(* IEC 61131-3 sources: plc-st-coding-agent/progress/evidence/f14_p1_20261111b/jobs/codex_deepseek-v4pro, 35 files *)

(* ---- public-easy-02.candidate_01.st ---- *)
FUNCTION_BLOCK DualWordEdgeDetector
VAR_INPUT
    value : DWORD;
END_VAR
VAR_OUTPUT
    hasChanged       : BOOL;
    hasRisingEdges   : BOOL;
    risingBits       : DWORD;
    noOfRisingBits   : USINT;
    hasFallingEdges  : BOOL;
    fallingBits      : DWORD;
    noOfFallingBits  : USINT;
END_VAR
VAR
    prevValue : DWORD;
    i : INT;
END_VAR

risingBits := value AND NOT prevValue;
fallingBits := NOT value AND prevValue;

hasRisingEdges := risingBits <> 0;
hasFallingEdges := fallingBits <> 0;
hasChanged := value <> prevValue;

noOfRisingBits := 0;
noOfFallingBits := 0;

FOR i := 0 TO 31 DO
    IF (risingBits AND SHL(DWORD#1, i)) <> 0 THEN
        noOfRisingBits := noOfRisingBits + 1;
    END_IF;

    IF (fallingBits AND SHL(DWORD#1, i)) <> 0 THEN
        noOfFallingBits := noOfFallingBits + 1;
    END_IF;
END_FOR;

prevValue := value;

(* ---- public-easy-02.candidate_02.st ---- *)
FUNCTION_BLOCK DualWordEdgeDetector
VAR_INPUT
    value : DWORD;
END_VAR
VAR_OUTPUT
    hasChanged       : BOOL;
    hasRisingEdges   : BOOL;
    risingBits       : DWORD;
    noOfRisingBits   : USINT;
    hasFallingEdges  : BOOL;
    fallingBits      : DWORD;
    noOfFallingBits  : USINT;
END_VAR
VAR
    prevValue : DWORD;
    i : INT;
END_VAR

risingBits := value AND (NOT prevValue);
fallingBits := (NOT value) AND prevValue;

hasRisingEdges := risingBits <> 0;
hasFallingEdges := fallingBits <> 0;
hasChanged := value <> prevValue;

noOfRisingBits := 0;
noOfFallingBits := 0;

FOR i := 0 TO 31 DO
    IF (risingBits AND SHL(DWORD#1, i)) <> 0 THEN
        noOfRisingBits := noOfRisingBits + 1;
    END_IF;

    IF (fallingBits AND SHL(DWORD#1, i)) <> 0 THEN
        noOfFallingBits := noOfFallingBits + 1;
    END_IF;
END_FOR;

prevValue := value;

END_FUNCTION_BLOCK

(* ---- public-easy-05.candidate_01.st ---- *)
FUNCTION_BLOCK WeldGapAlarm
VAR_INPUT
    Gap_Exceeded       : BOOL;
    Weld_E_Stop_NC     : BOOL;
    DebounceTime       : TIME;
END_VAR
VAR_OUTPUT
    Operator_Alert         : BOOL;
    Weld_Soft_Start_Active : BOOL;
END_VAR
VAR
    PowerUpTimer  : TON;
    GapTimer      : TON;
END_VAR

// 5-second power-up initialization inhibition
PowerUpTimer(IN := TRUE, PT := T#5S);
Weld_Soft_Start_Active := NOT PowerUpTimer.Q;

// Gap debounce only after initialization and while emergency stop is inactive
GapTimer(
    IN := Gap_Exceeded
          AND PowerUpTimer.Q
          AND Weld_E_Stop_NC,
    PT := DebounceTime
);

// Alarm only after full debounce, and emergency stop overrides immediately
Operator_Alert := GapTimer.Q AND Weld_E_Stop_NC;

(* ---- public-easy-05.candidate_02.st ---- *)
FUNCTION_BLOCK WeldGapAlarm
VAR_INPUT
    Gap_Exceeded       : BOOL;
    Weld_E_Stop_NC     : BOOL;
    DebounceTime       : TIME;
END_VAR
VAR_OUTPUT
    Operator_Alert         : BOOL;
    Weld_Soft_Start_Active : BOOL;
END_VAR
VAR
    PowerUpTimer  : TON;
    GapTimer      : TON;
END_VAR

PowerUpTimer(IN := TRUE, PT := T#5S);
Weld_Soft_Start_Active := NOT PowerUpTimer.Q;

GapTimer(
    IN := Gap_Exceeded
          AND PowerUpTimer.Q
          AND Weld_E_Stop_NC,
    PT := DebounceTime
);

Operator_Alert := GapTimer.Q AND Weld_E_Stop_NC;

END_FUNCTION_BLOCK

(* ---- public-easy-06.candidate_01.st ---- *)
FUNCTION_BLOCK AerationBlowerControl
VAR_INPUT
    DO_LOW : BOOL;
    AERATION_E_STOP_NC : BOOL;
END_VAR
VAR_OUTPUT
    BLOWER_RUN : BOOL;
    AERATION_BLOWER_CYCLE_COUNT : UINT;
END_VAR
VAR
    StartDelay : TON;
    BlowerRunPrev : BOOL := FALSE;
    InitDone : BOOL := FALSE;
END_VAR

IF NOT InitDone THEN
    StartDelay(IN := FALSE, PT := T#5s);
    BLOWER_RUN := FALSE;
    AERATION_BLOWER_CYCLE_COUNT := 0;
    BlowerRunPrev := FALSE;
    InitDone := TRUE;
END_IF;

StartDelay(IN := DO_LOW AND AERATION_E_STOP_NC, PT := T#5s);
BLOWER_RUN := StartDelay.Q;

IF BLOWER_RUN AND NOT BlowerRunPrev THEN
    AERATION_BLOWER_CYCLE_COUNT := AERATION_BLOWER_CYCLE_COUNT + 1;
END_IF;

BlowerRunPrev := BLOWER_RUN;
END_FUNCTION_BLOCK

(* ---- public-hard-01.candidate_01.st ---- *)
FUNCTION_BLOCK MaterialProportioningControl
VAR_INPUT
    estop            : BOOL;  (* FALSE = emergency stop active *)
    opeMode          : BOOL;  (* FALSE = manual, TRUE = automatic *)
    valveAStart      : BOOL;
    valveBStart      : BOOL;
    valveCStart      : BOOL;
    valveDStart      : BOOL;
    mixMotorStart    : BOOL;
    autoStart        : BOOL;
    processMode      : BOOL;  (* FALSE = no C, TRUE = use C until 100 cm *)
    levelSensor      : INT;   (* cm *)
    mixMotorComplete : BOOL;
END_VAR

VAR_OUTPUT
    valveARun   : BOOL;
    valveBRun   : BOOL;
    valveCRun   : BOOL;
    valveDRun   : BOOL;
    mixMotorRun : BOOL;
END_VAR

VAR
    valveAStart_RE      : BOOL;
    valveBStart_RE      : BOOL;
    valveCStart_RE      : BOOL;
    valveDStart_RE      : BOOL;
    mixMotorStart_RE    : BOOL;
    autoStart_RE        : BOOL;
    mixMotorComplete_RE : BOOL;
    modeChanged         : BOOL;

    valveAStart_prev      : BOOL;
    valveBStart_prev      : BOOL;
    valveCStart_prev      : BOOL;
    valveDStart_prev      : BOOL;
    mixMotorStart_prev    : BOOL;
    autoStart_prev        : BOOL;
    mixMotorComplete_prev : BOOL;
    opeMode_prev          : BOOL;

    manualValveA   : BOOL;
    manualValveB   : BOOL;
    manualValveC   : BOOL;
    manualValveD   : BOOL;
    manualMixMotor : BOOL;

    (* 0  = idle *)
    (* 10 = filling through valve A *)
    (* 20 = filling through valve B *)
    (* 30 = filling through valve C *)
    (* 40 = mixing *)
    (* 50 = discharging through valve D *)
    autoState : INT := 0;
END_VAR

(* Detect rising edges *)
valveAStart_RE      := valveAStart AND NOT valveAStart_prev;
valveBStart_RE      := valveBStart AND NOT valveBStart_prev;
valveCStart_RE      := valveCStart AND NOT valveCStart_prev;
valveDStart_RE      := valveDStart AND NOT valveDStart_prev;
mixMotorStart_RE    := mixMotorStart AND NOT mixMotorStart_prev;
autoStart_RE        := autoStart AND NOT autoStart_prev;
mixMotorComplete_RE := mixMotorComplete AND NOT mixMotorComplete_prev;
modeChanged         := opeMode <> opeMode_prev;

IF NOT estop THEN
    (* Emergency stop: stop everything and reset control states *)
    valveARun   := FALSE;
    valveBRun   := FALSE;
    valveCRun   := FALSE;
    valveDRun   := FALSE;
    mixMotorRun := FALSE;

    autoState      := 0;
    manualValveA   := FALSE;
    manualValveB   := FALSE;
    manualValveC   := FALSE;
    manualValveD   := FALSE;
    manualMixMotor := FALSE;

ELSIF modeChanged THEN
    (* Mode change: stop equipment and clear both control states *)
    valveARun   := FALSE;
    valveBRun   := FALSE;
    valveCRun   := FALSE;
    valveDRun   := FALSE;
    mixMotorRun := FALSE;

    autoState      := 0;
    manualValveA   := FALSE;
    manualValveB   := FALSE;
    manualValveC   := FALSE;
    manualValveD   := FALSE;
    manualMixMotor := FALSE;

ELSIF opeMode THEN
    (* Automatic mode *)

    IF autoStart_RE AND ((autoState = 0) OR (autoState = 50)) THEN
        autoState := 10;
    END_IF;

    CASE autoState OF
        10: (* Valve A is open; fill to 50 cm *)
            IF levelSensor >= 50 THEN
                autoState := 20;
            END_IF;

        20: (* Valve A closed, valve B open; fill to 80 cm *)
            IF levelSensor >= 80 THEN
                IF processMode THEN
                    autoState := 30;
                ELSE
                    autoState := 40;
                END_IF;
            END_IF;

        30: (* Valve C open; fill to 100 cm *)
            IF levelSensor >= 100 THEN
                autoState := 40;
            END_IF;

        40: (* Mixing motor running *)
            IF mixMotorComplete_RE THEN
                autoState := 50;
            END_IF;

        50: (* Valve D open; automatic process finished *)
            ;
    END_CASE;

    valveARun   := autoState = 10;
    valveBRun   := autoState = 20;
    valveCRun   := autoState = 30;
    valveDRun   := autoState = 50;
    mixMotorRun := autoState = 40;

ELSE
    (* Manual mode: each rising edge toggles the corresponding device *)
    valveARun   := manualValveA;
    valveBRun   := manualValveB;
    valveCRun   := manualValveC;
    valveDRun   := manualValveD;
    mixMotorRun := manualMixMotor;

    IF valveAStart_RE THEN
        manualValveA := NOT manualValveA;
    END_IF;

    IF valveBStart_RE THEN
        manualValveB := NOT manualValveB;
    END_IF;

    IF valveCStart_RE THEN
        manualValveC := NOT manualValveC;
    END_IF;

    IF valveDStart_RE THEN
        manualValveD := NOT manualValveD;
    END_IF;

    IF mixMotorStart_RE THEN
        manualMixMotor := NOT manualMixMotor;
    END_IF;
END_IF;

(* Store current input values for the next rising-edge detection *)
valveAStart_prev      := valveAStart;
valveBStart_prev      := valveBStart;
valveCStart_prev      := valveCStart;
valveDStart_prev      := valveDStart;
mixMotorStart_prev    := mixMotorStart;
autoStart_prev        := autoStart;
mixMotorComplete_prev := mixMotorComplete;
opeMode_prev          := opeMode;

(* ---- public-hard-01.candidate_02.st ---- *)
FUNCTION_BLOCK MaterialProportioningControl
VAR_INPUT
    estop            : BOOL;  (* FALSE: emergency stop triggered *)
    opeMode          : BOOL;  (* FALSE: manual, TRUE: automatic *)
    valveAStart      : BOOL;
    valveBStart      : BOOL;
    valveCStart      : BOOL;
    valveDStart      : BOOL;
    mixMotorStart    : BOOL;
    autoStart        : BOOL;
    processMode      : BOOL;
    levelSensor      : INT;   (* cm *)
    mixMotorComplete : BOOL;
END_VAR

VAR_OUTPUT
    valveARun   : BOOL;
    valveBRun   : BOOL;
    valveCRun   : BOOL;
    valveDRun   : BOOL;
    mixMotorRun : BOOL;
END_VAR

VAR
    valveAStart_RE      : BOOL;
    valveBStart_RE      : BOOL;
    valveCStart_RE      : BOOL;
    valveDStart_RE      : BOOL;
    mixMotorStart_RE    : BOOL;
    autoStart_RE        : BOOL;
    mixMotorComplete_RE : BOOL;
    modeChanged         : BOOL;

    valveAStart_prev      : BOOL;
    valveBStart_prev      : BOOL;
    valveCStart_prev      : BOOL;
    valveDStart_prev      : BOOL;
    mixMotorStart_prev    : BOOL;
    autoStart_prev        : BOOL;
    mixMotorComplete_prev : BOOL;
    opeMode_prev          : BOOL;

    manualValveA   : BOOL;
    manualValveB   : BOOL;
    manualValveC   : BOOL;
    manualValveD   : BOOL;
    manualMixMotor : BOOL;

    autoState : INT := 0; (* 0=idle,10=A,20=B,30=C,40=mix,50=discharge *)
END_VAR

(* Rising edge detection *)
valveAStart_RE      := valveAStart AND NOT valveAStart_prev;
valveBStart_RE      := valveBStart AND NOT valveBStart_prev;
valveCStart_RE      := valveCStart AND NOT valveCStart_prev;
valveDStart_RE      := valveDStart AND NOT valveDStart_prev;
mixMotorStart_RE    := mixMotorStart AND NOT mixMotorStart_prev;
autoStart_RE        := autoStart AND NOT autoStart_prev;
mixMotorComplete_RE := mixMotorComplete AND NOT mixMotorComplete_prev;
modeChanged         := opeMode <> opeMode_prev;

IF NOT estop THEN
    (* Emergency stop: stop all equipment and reset control states *)
    valveARun   := FALSE;
    valveBRun   := FALSE;
    valveCRun   := FALSE;
    valveDRun   := FALSE;
    mixMotorRun := FALSE;

    autoState      := 0;
    manualValveA   := FALSE;
    manualValveB   := FALSE;
    manualValveC   := FALSE;
    manualValveD   := FALSE;
    manualMixMotor := FALSE;

ELSIF modeChanged THEN
    (* Mode change: stop all equipment and clear both mode states *)
    valveARun   := FALSE;
    valveBRun   := FALSE;
    valveCRun   := FALSE;
    valveDRun   := FALSE;
    mixMotorRun := FALSE;

    autoState      := 0;
    manualValveA   := FALSE;
    manualValveB   := FALSE;
    manualValveC   := FALSE;
    manualValveD   := FALSE;
    manualMixMotor := FALSE;

ELSIF opeMode THEN
    (* Automatic mode *)
    IF autoStart_RE AND ((autoState = 0) OR (autoState = 50)) THEN
        autoState := 10;
    END_IF;

    CASE autoState OF
        10:
            IF levelSensor >= 50 THEN
                autoState := 20;
            END_IF;

        20:
            IF levelSensor >= 80 THEN
                IF processMode THEN
                    autoState := 30;
                ELSE
                    autoState := 40;
                END_IF;
            END_IF;

        30:
            IF levelSensor >= 100 THEN
                autoState := 40;
            END_IF;

        40:
            IF mixMotorComplete_RE THEN
                autoState := 50;
            END_IF;

        50:
            ; (* Valve D remains open; automatic process finished *)
    END_CASE;

    valveARun   := autoState = 10;
    valveBRun   := autoState = 20;
    valveCRun   := autoState = 30;
    valveDRun   := autoState = 50;
    mixMotorRun := autoState = 40;

ELSE
    (* Manual mode *)
    IF valveAStart_RE THEN
        manualValveA := NOT manualValveA;
    END_IF;

    IF valveBStart_RE THEN
        manualValveB := NOT manualValveB;
    END_IF;

    IF valveCStart_RE THEN
        manualValveC := NOT manualValveC;
    END_IF;

    IF valveDStart_RE THEN
        manualValveD := NOT manualValveD;
    END_IF;

    IF mixMotorStart_RE THEN
        manualMixMotor := NOT manualMixMotor;
    END_IF;

    valveARun   := manualValveA;
    valveBRun   := manualValveB;
    valveCRun   := manualValveC;
    valveDRun   := manualValveD;
    mixMotorRun := manualMixMotor;
END_IF;

(* Save current input states for next edge detection *)
valveAStart_prev      := valveAStart;
valveBStart_prev      := valveBStart;
valveCStart_prev      := valveCStart;
valveDStart_prev      := valveDStart;
mixMotorStart_prev    := mixMotorStart;
autoStart_prev        := autoStart;
mixMotorComplete_prev := mixMotorComplete;
opeMode_prev          := opeMode;

END_FUNCTION_BLOCK

(* ---- public-hard-05.candidate_01.st ---- *)
FUNCTION_BLOCK MechanicalArmControl
VAR_INPUT
    ManualMode        : BOOL;
    SingleStepMode    : BOOL;
    SingleCycleMode   : BOOL;
    ContinuousMode    : BOOL;
    EmergencyStop     : BOOL; (* FALSE: emergency stop triggered; TRUE: normal *)
    Start             : BOOL;
    DownButton        : BOOL;
    UpButton          : BOOL;
    LeftButton        : BOOL;
    RightButton       : BOOL;
    GripButton        : BOOL;
    ReleaseButton     : BOOL;
    DownLimitSwitch   : BOOL;
    UpLimitSwitch     : BOOL;
    LeftLimitSwitch   : BOOL;
    RightLimitSwitch  : BOOL;
    GripLimitSwitch   : BOOL;
    ReleaseLimitSwitch: BOOL;
END_VAR

VAR_OUTPUT
    MoveDown        : BOOL;
    MoveUp          : BOOL;
    MoveLeft        : BOOL;
    MoveRight       : BOOL;
    ActivateGrip    : BOOL;
    ActivateRelease : BOOL;
END_VAR

VAR
    StartPrev        : BOOL := FALSE;
    StartEdge        : BOOL := FALSE;
    StepActive       : BOOL := FALSE;
    StepIndex        : INT  := 0;
    SingleCycleState : INT  := 0;
    ContinuousState  : INT  := 0;
END_VAR

(* Rising edge of Start *)
StartEdge := Start AND NOT StartPrev;
StartPrev := Start;

(* Clear all commands first; emergency stop therefore disables all outputs. *)
MoveDown        := FALSE;
MoveUp          := FALSE;
MoveLeft        := FALSE;
MoveRight       := FALSE;
ActivateGrip    := FALSE;
ActivateRelease := FALSE;

IF NOT EmergencyStop THEN
    StartEdge := FALSE;

    StepActive       := FALSE;
    StepIndex        := 0;
    SingleCycleState := 0;
    ContinuousState  := 0;
ELSE
    (* ---------- Manual mode ---------- *)
    IF ManualMode THEN
        MoveDown        := DownButton    AND NOT DownLimitSwitch;
        MoveUp          := UpButton      AND NOT UpLimitSwitch;
        MoveLeft        := LeftButton    AND NOT LeftLimitSwitch;
        MoveRight       := RightButton   AND NOT RightLimitSwitch;
        ActivateGrip    := GripButton    AND NOT GripLimitSwitch;
        ActivateRelease := ReleaseButton AND NOT ReleaseLimitSwitch;
    END_IF;

    (* ---------- Single step mode ---------- *)
    IF SingleStepMode THEN
        IF StartEdge THEN
            StepIndex := StepIndex + 1;
            IF StepIndex > 8 THEN
                StepIndex := 1;
            END_IF;
            StepActive := TRUE;
        END_IF;

        IF StepActive THEN
            CASE StepIndex OF
                1: (* Down *)
                    IF DownLimitSwitch THEN
                        StepActive := FALSE;
                    ELSE
                        MoveDown := TRUE;
                    END_IF;
                2: (* Grip *)
                    IF GripLimitSwitch THEN
                        StepActive := FALSE;
                    ELSE
                        ActivateGrip := TRUE;
                    END_IF;
                3: (* Up *)
                    IF UpLimitSwitch THEN
                        StepActive := FALSE;
                    ELSE
                        MoveUp := TRUE;
                    END_IF;
                4: (* Right *)
                    IF RightLimitSwitch THEN
                        StepActive := FALSE;
                    ELSE
                        MoveRight := TRUE;
                    END_IF;
                5: (* Down *)
                    IF DownLimitSwitch THEN
                        StepActive := FALSE;
                    ELSE
                        MoveDown := TRUE;
                    END_IF;
                6: (* Release *)
                    IF ReleaseLimitSwitch THEN
                        StepActive := FALSE;
                    ELSE
                        ActivateRelease := TRUE;
                    END_IF;
                7: (* Up *)
                    IF UpLimitSwitch THEN
                        StepActive := FALSE;
                    ELSE
                        MoveUp := TRUE;
                    END_IF;
                8: (* Left *)
                    IF LeftLimitSwitch THEN
                        StepActive := FALSE;
                    ELSE
                        MoveLeft := TRUE;
                    END_IF;
            END_CASE;
        END_IF;
    ELSE
        StepActive := FALSE;
        StepIndex  := 0;
    END_IF;

    (* ---------- Single cycle mode ---------- *)
    IF SingleCycleMode THEN
        CASE SingleCycleState OF
            0: (* Idle, wait for Start *)
                IF StartEdge THEN
                    SingleCycleState := 1;
                END_IF;
            1: (* Down *)
                IF DownLimitSwitch THEN
                    SingleCycleState := 2;
                ELSE
                    MoveDown := TRUE;
                END_IF;
            2: (* Grip *)
                IF GripLimitSwitch THEN
                    SingleCycleState := 3;
                ELSE
                    ActivateGrip := TRUE;
                END_IF;
            3: (* Up *)
                IF UpLimitSwitch THEN
                    SingleCycleState := 4;
                ELSE
                    MoveUp := TRUE;
                END_IF;
            4: (* Right *)
                IF RightLimitSwitch THEN
                    SingleCycleState := 5;
                ELSE
                    MoveRight := TRUE;
                END_IF;
            5: (* Down *)
                IF DownLimitSwitch THEN
                    SingleCycleState := 6;
                ELSE
                    MoveDown := TRUE;
                END_IF;
            6: (* Release *)
                IF ReleaseLimitSwitch THEN
                    SingleCycleState := 7;
                ELSE
                    ActivateRelease := TRUE;
                END_IF;
            7: (* Up *)
                IF UpLimitSwitch THEN
                    SingleCycleState := 8;
                ELSE
                    MoveUp := TRUE;
                END_IF;
            8: (* Left *)
                IF LeftLimitSwitch THEN
                    SingleCycleState := 9;
                ELSE
                    MoveLeft := TRUE;
                END_IF;
            9: (* Completed; wait for next Start *)
                IF StartEdge THEN
                    SingleCycleState := 1;
                END_IF;
        END_CASE;
    ELSE
        SingleCycleState := 0;
    END_IF;

    (* ---------- Continuous mode ---------- *)
    IF ContinuousMode THEN
        CASE ContinuousState OF
            0: (* Idle, wait for Start *)
                IF StartEdge THEN
                    ContinuousState := 1;
                END_IF;
            1: (* Down *)
                IF DownLimitSwitch THEN
                    ContinuousState := 2;
                ELSE
                    MoveDown := TRUE;
                END_IF;
            2: (* Grip *)
                IF GripLimitSwitch THEN
                    ContinuousState := 3;
                ELSE
                    ActivateGrip := TRUE;
                END_IF;
            3: (* Up *)
                IF UpLimitSwitch THEN
                    ContinuousState := 4;
                ELSE
                    MoveUp := TRUE;
                END_IF;
            4: (* Right *)
                IF RightLimitSwitch THEN
                    ContinuousState := 5;
                ELSE
                    MoveRight := TRUE;
                END_IF;
            5: (* Down *)
                IF DownLimitSwitch THEN
                    ContinuousState := 6;
                ELSE
                    MoveDown := TRUE;
                END_IF;
            6: (* Release *)
                IF ReleaseLimitSwitch THEN
                    ContinuousState := 7;
                ELSE
                    ActivateRelease := TRUE;
                END_IF;
            7: (* Up *)
                IF UpLimitSwitch THEN
                    ContinuousState := 8;
                ELSE
                    MoveUp := TRUE;
                END_IF;
            8: (* Left, then immediately start the next cycle *)
                IF LeftLimitSwitch THEN
                    ContinuousState := 1;
                ELSE
                    MoveLeft := TRUE;
                END_IF;
        END_CASE;
    ELSE
        ContinuousState := 0;
    END_IF;
END_IF;

END_FUNCTION_BLOCK

(* ---- public-medium-01.candidate_01.st ---- *)
TYPE ST_Pump :
STRUCT
    priority  : INT;
    selection : BOOL;
    RunComd   : BOOL;
END_STRUCT
END_TYPE

FUNCTION_BLOCK FB_MultiPumpControl
VAR_INPUT
    mode  : BOOL; // FALSE: Manual, TRUE: Automatic
    start : BOOL; // Start selected pumps
    stop  : BOOL; // Stop all pumps
END_VAR
VAR_IN_OUT
    pumpGroup : ARRAY[1..5] OF ST_Pump;
END_VAR
VAR
    runActive   : BOOL := FALSE;
    selected    : ARRAY[1..5] OF BOOL;
    i           : INT;
    rank        : INT;
    bestIndex   : INT;
    bestPriority: INT;
END_VAR

IF stop THEN
    runActive := FALSE;
ELSIF start THEN
    runActive := TRUE;
END_IF;

FOR i := 1 TO 5 DO
    selected[i] := FALSE;
END_FOR;

IF runActive THEN
    IF mode THEN
        FOR rank := 1 TO 3 DO
            bestIndex := 0;
            bestPriority := 0;

            FOR i := 1 TO 5 DO
                IF NOT selected[i] THEN
                    IF (bestIndex = 0) OR (pumpGroup[i].priority > bestPriority) THEN
                        bestIndex := i;
                        bestPriority := pumpGroup[i].priority;
                    END_IF;
                END_IF;
            END_FOR;

            IF bestIndex <> 0 THEN
                selected[bestIndex] := TRUE;
            END_IF;
        END_FOR;
    ELSE
        FOR i := 1 TO 5 DO
            selected[i] := pumpGroup[i].selection;
        END_FOR;
    END_IF;
END_IF;

FOR i := 1 TO 5 DO
    pumpGroup[i].RunComd := selected[i] AND runActive;
END_FOR;

(* ---- public-medium-01.candidate_02.st ---- *)
TYPE ST_Pump :
STRUCT
    priority  : INT;
    selection : BOOL;
    RunComd   : BOOL;
END_STRUCT
END_TYPE

FUNCTION_BLOCK FB_MultiPumpControl
VAR_INPUT
    mode  : BOOL; // FALSE: Manual, TRUE: Automatic
    start : BOOL; // Start selected pumps
    stop  : BOOL; // Stop all pumps
END_VAR
VAR_IN_OUT
    pumpGroup : ARRAY[1..5] OF ST_Pump;
END_VAR
VAR
    runActive   : BOOL := FALSE;
    selected    : ARRAY[1..5] OF BOOL;
    i           : INT;
    rank        : INT;
    bestIndex   : INT;
    bestPriority: INT;
END_VAR

IF stop THEN
    runActive := FALSE;
ELSIF start THEN
    runActive := TRUE;
END_IF;

FOR i := 1 TO 5 DO
    selected[i] := FALSE;
END_FOR;

IF runActive THEN
    IF mode THEN
        FOR rank := 1 TO 3 DO
            bestIndex := 0;
            bestPriority := 0;

            FOR i := 1 TO 5 DO
                IF NOT selected[i] THEN
                    IF (bestIndex = 0) OR (pumpGroup[i].priority > bestPriority) THEN
                        bestIndex := i;
                        bestPriority := pumpGroup[i].priority;
                    END_IF;
                END_IF;
            END_FOR;

            IF bestIndex <> 0 THEN
                selected[bestIndex] := TRUE;
            END_IF;
        END_FOR;
    ELSE
        FOR i := 1 TO 5 DO
            selected[i] := pumpGroup[i].selection;
        END_FOR;
    END_IF;
END_IF;

FOR i := 1 TO 5 DO
    pumpGroup[i].RunComd := selected[i] AND runActive;
END_FOR;

END_FUNCTION_BLOCK

(* ---- public-medium-04.candidate_01.st ---- *)
FUNCTION_BLOCK FB_TemperatureControl
VAR_INPUT
    TemperatureSensorInput : REAL;
    SetTemperature : REAL;
END_VAR
VAR_OUTPUT
    CurrentTemperature : REAL;
    SetTempDisplay : REAL;
    HeaterStatus : BOOL;
    OverheatProtection : BOOL;
    HeaterOutput : BOOL;
END_VAR
VAR
    SensorFault : BOOL;
    HeaterCommand : BOOL;
    HeaterOnTimer : TON;
    CoolDownTimer : TON;
END_VAR

(* Display values *)
CurrentTemperature := TemperatureSensorInput;
SetTempDisplay := SetTemperature;

(* Sensor fault: valid measurement range is 0.0 to 100.0 *)
SensorFault := (TemperatureSensorInput < 0.0) OR (TemperatureSensorInput > 100.0);

(* Overheating protection remains active for at least 3 seconds *)
CoolDownTimer(IN := OverheatProtection, PT := T#3S);
IF CoolDownTimer.Q THEN
    OverheatProtection := FALSE;
END_IF;

(* Normal heater command *)
HeaterCommand := (NOT SensorFault)
                 AND (NOT OverheatProtection)
                 AND (TemperatureSensorInput < SetTemperature);

(* Heater running continuously for more than 5 seconds triggers protection *)
HeaterOnTimer(IN := HeaterCommand, PT := T#5S);
IF HeaterOnTimer.Q THEN
    OverheatProtection := TRUE;
END_IF;

(* Force heater off if protection is active, including the trigger moment *)
HeaterOutput := HeaterCommand AND (NOT OverheatProtection);

(* Heater status indication *)
HeaterStatus := HeaterOutput;

END_FUNCTION_BLOCK

(* ---- public-medium-06.candidate_01.st ---- *)
FUNCTION_BLOCK FB_SlabThicknessFaultMonitor
VAR_INPUT
    THICKNESS_FAULT        : BOOL;
    THICKNESS_SIGNAL_VALID : BOOL;
    CUTTING_RUN            : BOOL;
    FaultTimestamp         : DINT;
    CycleTime              : TIME; (* Must be positive *)
END_VAR
VAR_OUTPUT
    THICKNESS_ALARM        : BOOL;
    Slab_Fault_Counter     : UINT;
    Slab_Runtime_Accumulator : LTIME;
    Slab_Fault_History     : ARRAY[0..4] OF DINT; (* Read-only to callers *)
END_VAR
VAR
    Initialized    : BOOL;
    ValidFault     : BOOL;
    FaultRise      : R_TRIG;
    HoldTimer      : TON;
    HoldActive     : BOOL;
    HistoryStore   : ARRAY[0..4] OF DINT;
    i              : INT;
END_VAR

ValidFault := THICKNESS_SIGNAL_VALID AND THICKNESS_FAULT;

(* Power-up initialization *)
IF NOT Initialized THEN
    Slab_Fault_Counter := UINT#0;
    Slab_Runtime_Accumulator := LTIME#0S;

    FOR i := 0 TO 4 DO
        HistoryStore[i] := DINT#0;
    END_FOR;

    HoldActive := FALSE;
    HoldTimer(IN := FALSE, PT := T#500MS);
    Initialized := TRUE;
END_IF;

FaultRise(CLK := ValidFault);

IF NOT THICKNESS_SIGNAL_VALID THEN
    (* Signal invalid: alarm off, no holding, no fault records *)
    THICKNESS_ALARM := FALSE;
    HoldActive := FALSE;
    HoldTimer(IN := FALSE, PT := T#500MS);
ELSE
    IF FaultRise.Q THEN
        (* New valid thickness fault occurrence *)
        Slab_Fault_Counter := Slab_Fault_Counter + UINT#1;

        FOR i := 4 TO 1 BY -1 DO
            HistoryStore[i] := HistoryStore[i - 1];
        END_FOR;
        HistoryStore[0] := FaultTimestamp;

        (* Retrigger the minimum alarm hold *)
        HoldActive := FALSE;
    END_IF;

    HoldTimer(IN := HoldActive, PT := T#500MS);

    IF HoldTimer.Q THEN
        HoldActive := FALSE;
    END_IF;

    IF FaultRise.Q THEN
        HoldActive := TRUE;
    END_IF;

    THICKNESS_ALARM := THICKNESS_FAULT OR HoldActive;
END_IF;

(* Accumulate normal cutting runtime only under valid, fault-free running conditions *)
IF THICKNESS_SIGNAL_VALID
   AND CUTTING_RUN
   AND NOT THICKNESS_FAULT
   AND (CycleTime > T#0MS) THEN
    Slab_Runtime_Accumulator := Slab_Runtime_Accumulator + TIME_TO_LTIME(CycleTime);
END_IF;

(* Expose history as a copy; internal storage remains protected from direct caller changes *)
Slab_Fault_History := HistoryStore;

(* ---- public-medium-06.candidate_02.st ---- *)
FUNCTION_BLOCK FB_SlabThicknessFaultMonitor
VAR_INPUT
    THICKNESS_FAULT        : BOOL;
    THICKNESS_SIGNAL_VALID : BOOL;
    CUTTING_RUN            : BOOL;
    FaultTimestamp         : DINT;
    CycleTime              : TIME; (* Must be positive *)
END_VAR
VAR_OUTPUT
    THICKNESS_ALARM        : BOOL;
    Slab_Fault_Counter     : UINT;
    Slab_Runtime_Accumulator : LTIME;
    Slab_Fault_History     : ARRAY[0..4] OF DINT; (* Read-only to callers *)
END_VAR
VAR
    Initialized    : BOOL;
    ValidFault     : BOOL;
    FaultRise      : R_TRIG;
    HoldTimer      : TON;
    HoldActive     : BOOL;
    HistoryStore   : ARRAY[0..4] OF DINT;
    i              : INT;
END_VAR

ValidFault := THICKNESS_SIGNAL_VALID AND THICKNESS_FAULT;

(* Power-up initialization *)
IF NOT Initialized THEN
    Slab_Fault_Counter := UINT#0;
    Slab_Runtime_Accumulator := LTIME#0S;

    FOR i := 0 TO 4 DO
        HistoryStore[i] := DINT#0;
    END_FOR;

    HoldActive := FALSE;
    HoldTimer(IN := FALSE, PT := T#500MS);
    Initialized := TRUE;
END_IF;

FaultRise(CLK := ValidFault);

IF NOT THICKNESS_SIGNAL_VALID THEN
    (* Signal invalid: alarm off, no holding, no fault records *)
    THICKNESS_ALARM := FALSE;
    HoldActive := FALSE;
    HoldTimer(IN := FALSE, PT := T#500MS);
ELSE
    IF FaultRise.Q THEN
        (* New valid thickness fault occurrence *)
        Slab_Fault_Counter := Slab_Fault_Counter + UINT#1;

        FOR i := 4 TO 1 BY -1 DO
            HistoryStore[i] := HistoryStore[i - 1];
        END_FOR;
        HistoryStore[0] := FaultTimestamp;

        (* Retrigger the minimum alarm hold *)
        HoldActive := FALSE;
    END_IF;

    HoldTimer(IN := HoldActive, PT := T#500MS);

    IF HoldTimer.Q THEN
        HoldActive := FALSE;
    END_IF;

    IF FaultRise.Q THEN
        HoldActive := TRUE;
    END_IF;

    THICKNESS_ALARM := THICKNESS_FAULT OR HoldActive;
END_IF;

(* Accumulate normal cutting runtime only under valid, fault-free running conditions *)
IF THICKNESS_SIGNAL_VALID
   AND CUTTING_RUN
   AND NOT THICKNESS_FAULT
   AND (CycleTime > T#0MS) THEN
    Slab_Runtime_Accumulator := Slab_Runtime_Accumulator + TIME_TO_LTIME(CycleTime);
END_IF;

(* Expose history as a copy; internal storage remains protected from direct caller changes *)
Slab_Fault_History := HistoryStore;

END_FUNCTION_BLOCK

(* ---- public-medium-08.candidate_01.st ---- *)
FUNCTION_BLOCK IPv4Parser
VAR_INPUT
    ipText : STRING(254);
END_VAR

VAR_OUTPUT
    ipValue : UDINT;
END_VAR

VAR
    index        : DINT;
    textLen      : DINT;
    dotCount     : DINT;
    currentByte  : BYTE;
    segmentValue : UDINT;
    inSegment    : BOOL;
    segments     : ARRAY[1..4] OF UDINT;
    digitValue   : UDINT;
END_VAR

ipValue := 0;
textLen := LEN(ipText);

IF textLen = 0 THEN
    RETURN;
END_IF;

dotCount := 0;
segmentValue := 0;
inSegment := FALSE;

FOR index := 1 TO textLen DO
    currentByte := ipText[index];

    IF currentByte = 46 THEN
        IF NOT inSegment OR dotCount >= 3 THEN
            RETURN;
        END_IF;

        IF segmentValue > 255 THEN
            RETURN;
        END_IF;

        segments[dotCount + 1] := segmentValue;
        dotCount := dotCount + 1;
        segmentValue := 0;
        inSegment := FALSE;
    ELSIF currentByte >= 48 AND currentByte <= 57 THEN
        IF currentByte = 48 THEN
            digitValue := 0;
        ELSIF currentByte = 49 THEN
            digitValue := 1;
        ELSIF currentByte = 50 THEN
            digitValue := 2;
        ELSIF currentByte = 51 THEN
            digitValue := 3;
        ELSIF currentByte = 52 THEN
            digitValue := 4;
        ELSIF currentByte = 53 THEN
            digitValue := 5;
        ELSIF currentByte = 54 THEN
            digitValue := 6;
        ELSIF currentByte = 55 THEN
            digitValue := 7;
        ELSIF currentByte = 56 THEN
            digitValue := 8;
        ELSE
            digitValue := 9;
        END_IF;

        IF segmentValue > 255 THEN
            RETURN;
        END_IF;

        segmentValue := segmentValue * 10 + digitValue;

        IF segmentValue > 255 THEN
            RETURN;
        END_IF;

        inSegment := TRUE;
    ELSE
        RETURN;
    END_IF;
END_FOR;

IF NOT inSegment OR dotCount <> 3 THEN
    RETURN;
END_IF;

segments[4] := segmentValue;

ipValue := segments[1] * 16777216
         + segments[2] * 65536
         + segments[3] * 256
         + segments[4];

END_FUNCTION_BLOCK

(* ---- self-easy-01.candidate_01.st ---- *)
FUNCTION_BLOCK FB
VAR_INPUT
    enable    : BOOL;
    values    : ARRAY[1..8] OF INT;
    count     : INT;
    avgEnable : BOOL;
END_VAR
VAR_OUTPUT
    avgOut    : REAL;
END_VAR
VAR
    sumValue   : DINT;
    sampleCount: INT;
    i          : INT;
END_VAR

IF enable AND avgEnable AND (count > 0) THEN
    sampleCount := count;

    IF sampleCount > 8 THEN
        sampleCount := 8;
    END_IF;

    sumValue := 0;

    FOR i := 1 TO sampleCount BY 1 DO
        sumValue := sumValue + INT_TO_DINT(values[i]);
    END_FOR;

    avgOut := DINT_TO_REAL(sumValue) / INT_TO_REAL(sampleCount);
END_IF;

END_FUNCTION_BLOCK

(* ---- self-easy-02.candidate_01.st ---- *)
FUNCTION_BLOCK FB
VAR_INPUT
    tankLevel        : REAL;   // 储罐液位百分比 0..100
    outletFlow       : REAL;   // 出口流量 m³/h（预留观测，本题不参与逻辑）
    inletPermit      : BOOL;   // 进料许可
    resetBtn         : BOOL;   // 复位按钮，上升沿有效
END_VAR
VAR_OUTPUT
    pumpRun          : BOOL;   // 进料泵运行命令
    alarmHigh        : BOOL;   // 高液位报警，自保持
    alarmLow         : BOOL;   // 低液位报警，自保持
    outletValveOpen  : BOOL;   // 出口阀开命令
END_VAR
VAR
    prevAlarmHigh    : BOOL := FALSE;
    prevAlarmLow     : BOOL := FALSE;
    prevResetBtn     : BOOL := FALSE;
END_VAR

// 高液位报警：危险条件优先于复位沿
alarmHigh := (tankLevel >= 85.0)
             OR (prevAlarmHigh AND NOT (resetBtn AND NOT prevResetBtn));

// 低液位报警：危险条件优先于复位沿
alarmLow := (tankLevel <= 15.0)
            OR (prevAlarmLow AND NOT (resetBtn AND NOT prevResetBtn));

// 任一报警有效时禁止进料泵运行
pumpRun := inletPermit AND NOT alarmHigh AND NOT alarmLow;

// 低报警有效期间关闭出口阀，其余情况开启
outletValveOpen := NOT alarmLow;

// 保存本拍状态，供下一扫描周期使用
prevAlarmHigh := alarmHigh;
prevAlarmLow  := alarmLow;
prevResetBtn  := resetBtn;

END_FUNCTION_BLOCK

(* ---- self-hard-01.candidate_01.st ---- *)
FUNCTION_BLOCK FB
VAR_INPUT
    flowLow : BOOL;
    ackBtn : BOOL;
    sensorOK : BOOL;
END_VAR
VAR_OUTPUT
    alarmActive : BOOL;
    alarmAcked : BOOL;
    highHigh : BOOL;
END_VAR
VAR
    lastAck : BOOL;
    lastFlowLow : BOOL;
    lastAlarmActive : BOOL;
    lastAlarmAcked : BOOL;
    ackRise : BOOL;
    lastFlowAndAcked : BOOL;
    lastFlowActiveAcked : BOOL;
END_VAR

ackRise := ackBtn AND NOT lastAck;

lastFlowAndAcked := lastFlowLow AND lastAlarmAcked;
lastFlowActiveAcked := lastFlowLow AND lastAlarmActive AND lastAlarmAcked;

highHigh := NOT sensorOK;

alarmActive := flowLow OR (lastAlarmActive AND NOT ackRise AND NOT lastFlowAndAcked);
alarmAcked := alarmActive AND (NOT flowLow OR ackRise OR lastFlowActiveAcked);

lastAck := ackBtn;
lastFlowLow := flowLow;
lastAlarmActive := alarmActive;
lastAlarmAcked := alarmAcked;

END_FUNCTION_BLOCK

(* ---- self-hard-02.candidate_01.st ---- *)
FUNCTION_BLOCK FB
VAR_INPUT
    startBtn : BOOL;
    abortBtn : BOOL;
    setpoint : REAL;
    pv : REAL;
    maxDuration : INT;
END_VAR
VAR_OUTPUT
    elapsed : INT;
    phase : INT;
    timeout : BOOL;
END_VAR
VAR
    lastStartBtn : BOOL;
    startRising : BOOL;
    prevPhase : INT;
    prevElapsed : INT;
    prevTimeout : BOOL;
END_VAR

startRising := startBtn AND NOT lastStartBtn;
prevPhase := phase;
prevElapsed := elapsed;
prevTimeout := timeout;

IF abortBtn THEN
    phase := 9;
    elapsed := prevElapsed;
    timeout := prevTimeout;
ELSIF startRising THEN
    phase := 1;
    elapsed := 0;
    timeout := FALSE;
ELSIF (prevPhase = 1) OR (prevPhase = 2) THEN
    elapsed := prevElapsed + 1;

    IF maxDuration <= elapsed THEN
        timeout := TRUE;
        phase := 3;
    ELSE
        timeout := FALSE;

        IF (prevPhase = 2) OR (pv >= setpoint) THEN
            phase := 2;
        ELSE
            phase := 1;
        END_IF;
    END_IF;
ELSE
    phase := prevPhase;
    elapsed := prevElapsed;
    timeout := prevTimeout;
END_IF;

lastStartBtn := startBtn;
END_FUNCTION_BLOCK

(* ---- self-hard-03.candidate_01.st ---- *)
FUNCTION_BLOCK FB
VAR_INPUT
    pushEn : BOOL;
    pushItem : INT;
    popEn : BOOL;
END_VAR
VAR_IN_OUT
    fifo : ARRAY[1..8] OF INT;
END_VAR
VAR_OUTPUT
    count : INT := 0;
    full : BOOL := FALSE;
    empty : BOOL := TRUE;
    head : INT := 0;
END_VAR
VAR
    pushRise : BOOL;
    popRise : BOOL;
    pushPrev : BOOL := FALSE;
    popPrev : BOOL := FALSE;
    workingCount : INT;
    idx : INT;
END_VAR

pushRise := pushEn AND NOT pushPrev;
popRise := popEn AND NOT popPrev;

workingCount := count;

IF popRise AND (workingCount > 0) THEN
    IF workingCount > 1 THEN
        FOR idx := 1 TO workingCount - 1 DO
            fifo[idx] := fifo[idx + 1];
        END_FOR;
    END_IF;
    fifo[workingCount] := 0;
    workingCount := workingCount - 1;
END_IF;

IF pushRise AND (workingCount < 8) THEN
    fifo[workingCount + 1] := pushItem;
    workingCount := workingCount + 1;
END_IF;

count := workingCount;
full := (workingCount = 8);
empty := (workingCount = 0);

IF workingCount > 0 THEN
    head := fifo[1];
ELSE
    head := 0;
END_IF;

pushPrev := pushEn;
popPrev := popEn;
END_FUNCTION_BLOCK

(* ---- self-hard-04.candidate_01.st ---- *)
FUNCTION_BLOCK FB
VAR_INPUT
    demand : INT;
    runHours : ARRAY[1..5] OF LINT;
    rotated : BOOL;
END_VAR
VAR_OUTPUT
    leadPump : INT;
    lagPump : INT;
    runningCount : INT;
END_VAR
VAR
    previousLeadPump : INT := 0;
    previousLagPump : INT := 0;
    previousRunningCount : INT := 0;
    clippedDemand : INT;
    minimumPump : INT;
    minimumHours : LINT;
    lagCandidate : INT;
    pumpIndex : INT;
END_VAR

clippedDemand := demand;
IF clippedDemand < 0 THEN
    clippedDemand := 0;
ELSIF clippedDemand > 5 THEN
    clippedDemand := 5;
END_IF;

runningCount := clippedDemand;

IF clippedDemand <= 0 THEN
    leadPump := 0;
    lagPump := 0;
ELSE
    minimumHours := runHours[1];
    minimumPump := 1;
    FOR pumpIndex := 2 TO 5 DO
        IF (runHours[pumpIndex] < minimumHours) OR
           ((runHours[pumpIndex] = minimumHours) AND (pumpIndex < minimumPump)) THEN
            minimumHours := runHours[pumpIndex];
            minimumPump := pumpIndex;
        END_IF;
    END_FOR;

    IF (previousLeadPump < 1) OR (previousLeadPump > 5) THEN
        leadPump := minimumPump;
    ELSIF rotated AND
          (previousLeadPump >= 1) AND
          (previousLeadPump <= 5) AND
          (runHours[previousLeadPump] - minimumHours > 50) THEN
        leadPump := minimumPump;
    ELSE
        leadPump := previousLeadPump;
    END_IF;

    IF clippedDemand >= 2 THEN
        IF (leadPump <> previousLeadPump) OR (runningCount > previousRunningCount) THEN
            lagCandidate := 0;
            FOR pumpIndex := 1 TO 5 DO
                IF pumpIndex <> leadPump THEN
                    IF lagCandidate = 0 THEN
                        lagCandidate := pumpIndex;
                    ELSIF (runHours[pumpIndex] < runHours[lagCandidate]) OR
                          ((runHours[pumpIndex] = runHours[lagCandidate]) AND
                           (pumpIndex < lagCandidate)) THEN
                        lagCandidate := pumpIndex;
                    END_IF;
                END_IF;
            END_FOR;
            lagPump := lagCandidate;
        ELSE
            lagPump := previousLagPump;
        END_IF;
    ELSE
        lagPump := 0;
    END_IF;
END_IF;

previousLeadPump := leadPump;
previousLagPump := lagPump;
previousRunningCount := runningCount;
END_FUNCTION_BLOCK

(* ---- self-hard-05.candidate_01.st ---- *)
FUNCTION_BLOCK FB
VAR_INPUT
    runRequest : BOOL;
    flameOK : BOOL;
    o2Valid : BOOL;
    o2PV : REAL;
    baseAir : REAL;
    resetBtn : BOOL;
END_VAR
VAR_OUTPUT
    fuelPermit : BOOL;
    trimEnable : BOOL;
    airTrim : REAL;
    airCommand : REAL;
    tripLatched : BOOL;
    o2Fault : BOOL;
END_VAR
VAR
    tripMemory : BOOL;
    resetPrev : BOOL;
    resetRising : BOOL;
END_VAR

resetRising := resetBtn AND NOT resetPrev;

tripMemory := (runRequest AND NOT flameOK)
              OR (tripMemory AND NOT (resetRising AND NOT runRequest AND NOT flameOK));
tripLatched := tripMemory;

fuelPermit := runRequest AND flameOK AND NOT tripLatched;

o2Fault := NOT o2Valid OR o2PV < 0.0 OR o2PV > 21.0;

trimEnable := fuelPermit AND NOT o2Fault;

IF trimEnable THEN
    airTrim := 2.0 * (2.0 - o2PV);
    IF airTrim > 10.0 THEN
        airTrim := 10.0;
    END_IF;
    IF airTrim < -10.0 THEN
        airTrim := -10.0;
    END_IF;
ELSE
    airTrim := 0.0;
END_IF;

IF fuelPermit THEN
    airCommand := baseAir + airTrim;
    IF airCommand > 100.0 THEN
        airCommand := 100.0;
    END_IF;
    IF airCommand < 0.0 THEN
        airCommand := 0.0;
    END_IF;
ELSE
    airCommand := 0.0;
END_IF;

resetPrev := resetBtn;

(* ---- self-hard-05.candidate_02.st ---- *)
FUNCTION_BLOCK FB
VAR_INPUT
    runRequest : BOOL;
    flameOK : BOOL;
    o2Valid : BOOL;
    o2PV : REAL;
    baseAir : REAL;
    resetBtn : BOOL;
END_VAR
VAR_OUTPUT
    fuelPermit : BOOL;
    trimEnable : BOOL;
    airTrim : REAL;
    airCommand : REAL;
    tripLatched : BOOL;
    o2Fault : BOOL;
END_VAR
VAR
    tripMemory : BOOL;
    resetPrev : BOOL;
    resetRising : BOOL;
END_VAR

resetRising := resetBtn AND NOT resetPrev;

tripMemory := (runRequest AND NOT flameOK)
              OR (tripMemory AND NOT (resetRising AND NOT runRequest AND NOT flameOK));
tripLatched := tripMemory;

fuelPermit := runRequest AND flameOK AND NOT tripLatched;

o2Fault := NOT o2Valid OR o2PV < 0.0 OR o2PV > 21.0;

trimEnable := fuelPermit AND NOT o2Fault;

IF trimEnable THEN
    airTrim := 2.0 * (2.0 - o2PV);

    IF airTrim > 10.0 THEN
        airTrim := 10.0;
    END_IF;

    IF airTrim < -10.0 THEN
        airTrim := -10.0;
    END_IF;
ELSE
    airTrim := 0.0;
END_IF;

IF fuelPermit THEN
    airCommand := baseAir + airTrim;

    IF airCommand > 100.0 THEN
        airCommand := 100.0;
    END_IF;

    IF airCommand < 0.0 THEN
        airCommand := 0.0;
    END_IF;
ELSE
    airCommand := 0.0;
END_IF;

resetPrev := resetBtn;

END_FUNCTION_BLOCK

(* ---- self-hard-06.candidate_01.st ---- *)
FUNCTION_BLOCK FB
VAR_INPUT
    runRequest : BOOL;
    pressure : REAL;
    pressureValid : BOOL;
    fuelFlow : REAL;
    steamFlow : REAL;
    outletCmd : INT;
    outletFeedback : INT;
    resetBtn : BOOL;
END_VAR
VAR_OUTPUT
    tripLatched : BOOL;
    fuelPermit : BOOL;
    currentCauseMask : WORD;
    latchedCauseMask : WORD;
    diagnosticActive : BOOL;
END_VAR
VAR
    resetPrev : BOOL := FALSE;
    resetRising : BOOL;
    resetAllowed : BOOL;
    tripPending : BOOL;
    overpressureActive : BOOL;
    valveStuckActive : BOOL;
    stuckCounter : INT := 0;
END_VAR

resetRising := resetBtn AND NOT resetPrev;

overpressureActive := runRequest AND pressureValid AND (pressure >= 4500.0);

IF overpressureActive AND (outletCmd >= 50) AND (outletFeedback <= 10) THEN
    IF stuckCounter < 3 THEN
        stuckCounter := stuckCounter + 1;
    END_IF;
ELSE
    stuckCounter := 0;
END_IF;

valveStuckActive := stuckCounter >= 3;

currentCauseMask := WORD#0;

IF runRequest AND NOT pressureValid THEN
    currentCauseMask := WORD#1;
ELSIF overpressureActive THEN
    IF valveStuckActive THEN
        currentCauseMask := currentCauseMask OR WORD#2;
    END_IF;

    IF (fuelFlow >= 4.0) AND (steamFlow <= 10.0) THEN
        currentCauseMask := currentCauseMask OR WORD#4;
    END_IF;

    IF currentCauseMask = WORD#0 THEN
        currentCauseMask := WORD#8;
    END_IF;
END_IF;

resetAllowed := resetRising AND NOT runRequest AND pressureValid AND (pressure <= 4200.0);
tripPending := runRequest AND ((NOT pressureValid) OR (pressure >= 4500.0));

IF resetAllowed THEN
    tripLatched := FALSE;
ELSE
    tripLatched := tripLatched OR tripPending;
END_IF;

fuelPermit := runRequest AND NOT tripLatched;
diagnosticActive := currentCauseMask <> WORD#0;

IF tripLatched THEN
    latchedCauseMask := latchedCauseMask OR currentCauseMask;
ELSE
    latchedCauseMask := WORD#0;
END_IF;

resetPrev := resetBtn;
END_FUNCTION_BLOCK

(* ---- self-hard-07.candidate_01.st ---- *)
FUNCTION_BLOCK FB
VAR_INPUT
    mode : INT;
    resetBtn : BOOL;
    scanSeconds : REAL;
    tempSP : REAL;
    tempPV : REAL;
    flowPV : REAL;
    manualFlowSP : REAL;
    manualValve : REAL;
END_VAR

VAR_OUTPUT
    flowSP : REAL;
    valveCommand : REAL;
    fault : BOOL;
    normalMode : BOOL;
END_VAR

VAR
    firstScan : BOOL := TRUE;
    prevMode : INT := 0;
    prevResetBtn : BOOL := FALSE;
    prevFlowSP : REAL := 0.0;
    prevValveCommand : REAL := 0.0;
    prevET : REAL := 0.0;
    prevEF : REAL := 0.0;
    resetRising : BOOL;
    modeChanged : BOOL;
    eT : REAL;
    eF : REAL;
END_VAR

    fault := (mode < 0) OR (mode > 2) OR (scanSeconds <= 0.0) OR (scanSeconds > 10.0);
    resetRising := resetBtn AND NOT prevResetBtn;
    modeChanged := (NOT firstScan) AND (mode <> prevMode);
    normalMode := (NOT firstScan) AND (mode = prevMode) AND (NOT fault) AND (NOT resetRising);

    eT := tempSP - tempPV;

    IF fault THEN
        flowSP := manualFlowSP;
        valveCommand := manualValve;
    ELSIF firstScan THEN
        flowSP := manualFlowSP;
        valveCommand := manualValve;
    ELSIF resetRising THEN
        flowSP := manualFlowSP;
        valveCommand := manualValve;
    ELSIF modeChanged THEN
        IF mode = 2 THEN
            flowSP := prevFlowSP;
            valveCommand := prevValveCommand;
        ELSE
            flowSP := manualFlowSP;
            valveCommand := prevValveCommand;
        END_IF;
    ELSE
        CASE mode OF
            0:
                flowSP := manualFlowSP;
                valveCommand := manualValve;

            1:
                flowSP := manualFlowSP;
                eF := flowSP - flowPV;
                valveCommand := LIMIT(0.0,
                    2.0 * eF + ((prevValveCommand - 2.0 * prevEF) + 0.5 * eF * scanSeconds),
                    100.0);

            2:
                flowSP := LIMIT(0.0,
                    1.0 * eT + ((prevFlowSP - 1.0 * prevET) + 0.2 * eT * scanSeconds),
                    50.0);
                eF := flowSP - flowPV;
                valveCommand := LIMIT(0.0,
                    2.0 * eF + ((prevValveCommand - 2.0 * prevEF) + 0.5 * eF * scanSeconds),
                    100.0);

            ELSE
                flowSP := manualFlowSP;
                valveCommand := manualValve;
        END_CASE;
    END_IF;

    prevResetBtn := resetBtn;
    prevMode := mode;
    prevFlowSP := flowSP;
    prevValveCommand := valveCommand;
    prevET := eT;
    prevEF := flowSP - flowPV;
    firstScan := FALSE;
END_FUNCTION_BLOCK

(* ---- self-medium-01.candidate_01.st ---- *)
FUNCTION_BLOCK FB
VAR_INPUT
    recipe : ARRAY[1..8] OF ST_Recipe;
    selSlot : INT;
    loadCmd : BOOL;
    running : BOOL;
END_VAR
VAR_OUTPUT
    valid : BOOL;
    loadedID : INT;
END_VAR
VAR
    previousLoadCmd : BOOL := FALSE;
    previousValid : BOOL := FALSE;
    previousLoadedID : INT := 0;
    loadEdge : BOOL;
    slotInRange : BOOL;
    slotNonEmpty : BOOL;
    ratioInRange : BOOL;
    temperatureInRange : BOOL;
END_VAR

loadEdge := loadCmd AND NOT previousLoadCmd;

loadedID := previousLoadedID;
valid := previousValid;

IF loadEdge AND NOT running THEN
    slotInRange := (selSlot >= 1) AND (selSlot <= 8);

    IF slotInRange THEN
        slotNonEmpty := recipe[selSlot].recipeID <> 0;
        ratioInRange := (recipe[selSlot].totalRatio >= 99.0)
                        AND (recipe[selSlot].totalRatio <= 101.0);
        temperatureInRange := (recipe[selSlot].temperature >= 30.0)
                              AND (recipe[selSlot].temperature <= 180.0);

        IF slotNonEmpty AND ratioInRange AND temperatureInRange THEN
            valid := TRUE;
            loadedID := recipe[selSlot].recipeID;
        ELSE
            valid := FALSE;
            loadedID := 0;
        END_IF;
    ELSE
        valid := FALSE;
        loadedID := 0;
    END_IF;
END_IF;

previousLoadCmd := loadCmd;
previousValid := valid;
previousLoadedID := loadedID;

(* ---- self-medium-01.candidate_02.st ---- *)
TYPE ST_Recipe :
STRUCT
    recipeID : INT;
    totalRatio : REAL;
    temperature : REAL;
END_STRUCT
END_TYPE

FUNCTION_BLOCK FB
VAR_INPUT
    recipe : ARRAY[1..8] OF ST_Recipe;
    selSlot : INT;
    loadCmd : BOOL;
    running : BOOL;
END_VAR
VAR_OUTPUT
    valid : BOOL;
    loadedID : INT;
END_VAR
VAR
    previousLoadCmd : BOOL := FALSE;
    previousValid : BOOL := FALSE;
    previousLoadedID : INT := 0;
    loadEdge : BOOL;
    slotInRange : BOOL;
    slotNonEmpty : BOOL;
    ratioInRange : BOOL;
    temperatureInRange : BOOL;
END_VAR

loadEdge := loadCmd AND NOT previousLoadCmd;

loadedID := previousLoadedID;
valid := previousValid;

IF loadEdge AND NOT running THEN
    slotInRange := (selSlot >= 1) AND (selSlot <= 8);

    IF slotInRange THEN
        slotNonEmpty := recipe[selSlot].recipeID <> 0;
        ratioInRange := (recipe[selSlot].totalRatio >= 99.0)
                        AND (recipe[selSlot].totalRatio <= 101.0);
        temperatureInRange := (recipe[selSlot].temperature >= 30.0)
                              AND (recipe[selSlot].temperature <= 180.0);

        IF slotNonEmpty AND ratioInRange AND temperatureInRange THEN
            valid := TRUE;
            loadedID := recipe[selSlot].recipeID;
        ELSE
            valid := FALSE;
            loadedID := 0;
        END_IF;
    ELSE
        valid := FALSE;
        loadedID := 0;
    END_IF;
END_IF;

previousLoadCmd := loadCmd;
previousValid := valid;
previousLoadedID := loadedID;

END_FUNCTION_BLOCK

(* ---- self-medium-02.candidate_01.st ---- *)
FUNCTION_BLOCK FB
VAR_INPUT
    enable : BOOL;
    rawValue : REAL;
END_VAR
VAR_OUTPUT
    filteredValue : REAL;
    windowFull : BOOL;
    sampleCount : INT;
END_VAR
VAR
    buffer : ARRAY[0..7] OF REAL;
    writeIndex : INT := 0;
    validCount : INT := 0;
    sum : REAL;
    loopIndex : INT;
END_VAR

IF enable THEN
    buffer[writeIndex] := rawValue;
    writeIndex := (writeIndex + 1) MOD 8;

    IF validCount < 8 THEN
        validCount := validCount + 1;
    END_IF;

    IF validCount = 1 THEN
        filteredValue := rawValue;
    ELSIF validCount = 2 THEN
        filteredValue := (buffer[0] + buffer[1]) / 2.0;
    ELSE
        sum := 0.0;
        FOR loopIndex := 0 TO validCount - 1 DO
            sum := sum + buffer[loopIndex];
        END_FOR;
        filteredValue := sum / INT_TO_REAL(validCount);
    END_IF;

    sampleCount := validCount;
    windowFull := validCount >= 8;
ELSE
    FOR loopIndex := 0 TO 7 DO
        buffer[loopIndex] := 0.0;
    END_FOR;

    writeIndex := 0;
    validCount := 0;
    sampleCount := 0;
    windowFull := FALSE;
END_IF

(* ---- self-medium-02.candidate_02.st ---- *)
FUNCTION_BLOCK FB
VAR_INPUT
    enable : BOOL;
    rawValue : REAL;
END_VAR
VAR_OUTPUT
    filteredValue : REAL;
    windowFull : BOOL;
    sampleCount : INT;
END_VAR
VAR
    buffer : ARRAY[0..7] OF REAL;
    writeIndex : INT := 0;
    validCount : INT := 0;
    sum : REAL;
    loopIndex : INT;
END_VAR

IF enable THEN
    buffer[writeIndex] := rawValue;
    writeIndex := (writeIndex + 1) MOD 8;

    IF validCount < 8 THEN
        validCount := validCount + 1;
    END_IF;

    IF validCount = 1 THEN
        filteredValue := rawValue;
    ELSIF validCount = 2 THEN
        filteredValue := (buffer[0] + buffer[1]) / 2.0;
    ELSE
        sum := 0.0;
        FOR loopIndex := 0 TO validCount - 1 DO
            sum := sum + buffer[loopIndex];
        END_FOR;
        filteredValue := sum / INT_TO_REAL(validCount);
    END_IF;

    sampleCount := validCount;
    windowFull := validCount >= 8;
ELSE
    FOR loopIndex := 0 TO 7 DO
        buffer[loopIndex] := 0.0;
    END_FOR;

    writeIndex := 0;
    validCount := 0;
    sampleCount := 0;
    windowFull := FALSE;
END_IF
END_FUNCTION_BLOCK

(* ---- self-medium-03.candidate_01.st ---- *)
FUNCTION_BLOCK FB
VAR_INPUT
    openBtn    : BOOL;
    closeBtn   : BOOL;
    openLimit  : BOOL;
    closeLimit : BOOL;
    obstacle   : BOOL;
END_VAR
VAR_OUTPUT
    motorUp    : BOOL;
    motorDown  : BOOL;
    errorFlag  : BOOL;
END_VAR
VAR
    state         : INT := 0; (* 0=IDLE, 1=OPENING, 2=CLOSING, 3=FAULT *)
    prevOpenBtn   : BOOL := FALSE;
    prevCloseBtn  : BOOL := FALSE;
    prevObstacle  : BOOL := FALSE;
    prevMotorUp   : BOOL := FALSE;
    prevMotorDown : BOOL := FALSE;
    prevErrorFlag : BOOL := FALSE;
END_VAR

VAR
    openRising  : BOOL;
    closeRising : BOOL;
    comboRising : BOOL;
END_VAR

openRising  := openBtn AND NOT prevOpenBtn;
closeRising := closeBtn AND NOT prevCloseBtn;
comboRising := (openBtn AND closeBtn) AND NOT (prevOpenBtn AND prevCloseBtn);

IF obstacle THEN
    state := 3;
    motorUp := FALSE;
    motorDown := FALSE;
    errorFlag := TRUE;
ELSIF state = 3 THEN
    motorUp := FALSE;
    motorDown := FALSE;
    IF comboRising THEN
        state := 0;
        errorFlag := FALSE;
    ELSE
        errorFlag := TRUE;
    END_IF;
ELSIF state = 1 THEN
    errorFlag := FALSE;
    motorDown := FALSE;
    IF openLimit THEN
        motorUp := FALSE;
        state := 0;
    ELSE
        motorUp := TRUE;
    END_IF;
ELSIF state = 2 THEN
    errorFlag := FALSE;
    motorUp := FALSE;
    IF closeLimit THEN
        motorDown := FALSE;
        state := 0;
    ELSE
        motorDown := TRUE;
    END_IF;
ELSE (* state = 0: IDLE *)
    motorUp := FALSE;
    motorDown := FALSE;
    errorFlag := FALSE;

    IF openRising AND NOT closeBtn AND NOT openLimit THEN
        motorUp := TRUE;
        state := 1;
    ELSIF closeRising AND NOT openBtn AND NOT closeLimit THEN
        motorDown := TRUE;
        state := 2;
    END_IF;
END_IF;

prevOpenBtn   := openBtn;
prevCloseBtn  := closeBtn;
prevObstacle  := obstacle;
prevMotorUp   := motorUp;
prevMotorDown := motorDown;
prevErrorFlag := errorFlag;
END_FUNCTION_BLOCK

(* ---- self-medium-04.candidate_01.st ---- *)
FUNCTION_BLOCK FB
VAR_INPUT
    startBtn : BOOL;
    resetBtn : BOOL;
    doneSensor : BOOL;
    targetVol : REAL;
    flowVol : REAL;
END_VAR
VAR_OUTPUT
    valveOpen : BOOL;
    fillsToday : INT;
END_VAR
VAR
    prevStartBtn : BOOL;
    prevResetBtn : BOOL;
    prevValveOpen : BOOL;
    bottleVol : REAL;
    pendingConfirm : BOOL;
    valveState : BOOL;
    fillCount : INT;
END_VAR

IF resetBtn AND NOT prevResetBtn THEN
    fillCount := 0;
    bottleVol := 0.0;
    valveState := FALSE;
    pendingConfirm := FALSE;
ELSE
    IF startBtn AND NOT prevStartBtn THEN
        IF NOT prevValveOpen THEN
            pendingConfirm := FALSE;
            bottleVol := 0.0;
            valveState := TRUE;
        END_IF;
    END_IF;

    IF valveState THEN
        bottleVol := bottleVol + flowVol;
        IF bottleVol >= targetVol THEN
            valveState := FALSE;
            pendingConfirm := TRUE;
        END_IF;
    END_IF;

    IF doneSensor AND pendingConfirm AND NOT valveState THEN
        IF fillCount < 32767 THEN
            fillCount := fillCount + 1;
        END_IF;
        pendingConfirm := FALSE;
    END_IF;
END_IF;

valveOpen := valveState;
fillsToday := fillCount;

prevStartBtn := startBtn;
prevResetBtn := resetBtn;
prevValveOpen := valveState;

(* ---- self-medium-04.candidate_02.st ---- *)
FUNCTION_BLOCK FB
VAR_INPUT
    startBtn : BOOL;
    resetBtn : BOOL;
    doneSensor : BOOL;
    targetVol : REAL;
    flowVol : REAL;
END_VAR
VAR_OUTPUT
    valveOpen : BOOL;
    fillsToday : INT;
END_VAR
VAR
    prevStartBtn : BOOL;
    prevResetBtn : BOOL;
    prevValveOpen : BOOL;
    bottleVol : REAL;
    pendingConfirm : BOOL;
    valveState : BOOL;
    fillCount : INT;
END_VAR

IF resetBtn AND NOT prevResetBtn THEN
    fillCount := 0;
    bottleVol := 0.0;
    valveState := FALSE;
    pendingConfirm := FALSE;
ELSE
    IF startBtn AND NOT prevStartBtn THEN
        IF NOT prevValveOpen THEN
            pendingConfirm := FALSE;
            bottleVol := 0.0;
            valveState := TRUE;
        END_IF;
    END_IF;

    IF valveState THEN
        bottleVol := bottleVol + flowVol;
        IF bottleVol >= targetVol THEN
            valveState := FALSE;
            pendingConfirm := TRUE;
        END_IF;
    END_IF;

    IF doneSensor AND pendingConfirm AND NOT valveState THEN
        IF fillCount < 32767 THEN
            fillCount := fillCount + 1;
        END_IF;
        pendingConfirm := FALSE;
    END_IF;
END_IF;

valveOpen := valveState;
fillsToday := fillCount;

prevStartBtn := startBtn;
prevResetBtn := resetBtn;
prevValveOpen := valveState;

END_FUNCTION_BLOCK

(* ---- self-medium-05.candidate_01.st ---- *)
FUNCTION_BLOCK FB
VAR_INPUT
    enable : BOOL;
    resetBtn : BOOL;
    scanSeconds : LREAL;
    steamFlow : LREAL;
    fuelFlow : LREAL;
    steamTemp : LREAL;
    steamPressure : LREAL;
END_VAR
VAR_OUTPUT
    qualified : BOOL;
    dataFault : BOOL;
    qualifiedTon : LREAL;
    fuelTon : LREAL;
    revenue : LREAL;
    cost : LREAL;
    netProfit : LREAL;
END_VAR
VAR
    resetBtnPrev : BOOL;
END_VAR

qualified := (steamTemp >= 447.0)
             AND (steamTemp <= 453.0)
             AND (steamPressure >= 3750.0)
             AND (steamPressure <= 3850.0);

dataFault := (scanSeconds <= 0.0)
             OR (scanSeconds > 10.0)
             OR (steamFlow < 0.0)
             OR (steamFlow > 90.0)
             OR (fuelFlow < 0.0)
             OR (fuelFlow > 6.0);

IF resetBtn AND NOT resetBtnPrev THEN
    qualifiedTon := 0.0;
    fuelTon := 0.0;
ELSIF dataFault THEN
    qualifiedTon := qualifiedTon;
    fuelTon := fuelTon;
ELSIF enable THEN
    fuelTon := fuelTon + fuelFlow * scanSeconds / 1000.0;

    IF qualified THEN
        qualifiedTon := qualifiedTon + steamFlow * scanSeconds / 1000.0;
    END_IF;
ELSIF NOT enable THEN
    qualifiedTon := qualifiedTon;
    fuelTon := fuelTon;
END_IF;

revenue := qualifiedTon * 280.0;
cost := fuelTon * 1500.0;
netProfit := revenue - cost;

resetBtnPrev := resetBtn;

(* ---- self-medium-05.candidate_02.st ---- *)
FUNCTION_BLOCK FB
VAR_INPUT
    enable : BOOL;
    resetBtn : BOOL;
    scanSeconds : LREAL;
    steamFlow : LREAL;
    fuelFlow : LREAL;
    steamTemp : LREAL;
    steamPressure : LREAL;
END_VAR
VAR_OUTPUT
    qualified : BOOL;
    dataFault : BOOL;
    qualifiedTon : LREAL;
    fuelTon : LREAL;
    revenue : LREAL;
    cost : LREAL;
    netProfit : LREAL;
END_VAR
VAR
    resetBtnPrev : BOOL := FALSE;
    qualifiedAcc : LREAL := 0.0;
    fuelAcc : LREAL := 0.0;
END_VAR

qualified := (steamTemp >= 447.0)
             AND (steamTemp <= 453.0)
             AND (steamPressure >= 3750.0)
             AND (steamPressure <= 3850.0);

dataFault := (scanSeconds <= 0.0)
             OR (scanSeconds > 10.0)
             OR (steamFlow < 0.0)
             OR (steamFlow > 90.0)
             OR (fuelFlow < 0.0)
             OR (fuelFlow > 6.0);

IF resetBtn AND NOT resetBtnPrev THEN
    qualifiedAcc := 0.0;
    fuelAcc := 0.0;
ELSE
    IF enable AND NOT dataFault THEN
        fuelAcc := fuelAcc + fuelFlow * scanSeconds / 1000.0;

        IF qualified THEN
            qualifiedAcc := qualifiedAcc + steamFlow * scanSeconds / 1000.0;
        END_IF;
    END_IF;
END_IF;

qualifiedTon := qualifiedAcc;
fuelTon := fuelAcc;

revenue := qualifiedTon * 280.0;
cost := fuelTon * 1500.0;
netProfit := revenue - cost;

resetBtnPrev := resetBtn;

END_FUNCTION_BLOCK

(* ---- public-easy-01.candidate_01.st ---- *)
PROGRAM FillingLineControl
VAR_INPUT
    bottleSensor : BOOL;
    cleaningConfirmButton : BOOL;
    fillingConfirmButton : BOOL;
    cappingConfirmButton : BOOL;
    packingConfirmButton : BOOL;
    finishedButton : BOOL;
END_VAR
VAR_OUTPUT
    Pump_Motor : BOOL;
    Filling_Valve : BOOL;
    Capping_Machine : BOOL;
    Packing_Machine : BOOL;
    Completion_Light : BOOL;
END_VAR
VAR
    State : INT := 0;
    bottleSensorR : R_TRIG;
    cleaningConfirmR : R_TRIG;
    fillingConfirmR : R_TRIG;
    cappingConfirmR : R_TRIG;
    packingConfirmR : R_TRIG;
    finishedR : R_TRIG;
END_VAR

bottleSensorR(CLK := bottleSensor);
cleaningConfirmR(CLK := cleaningConfirmButton);
fillingConfirmR(CLK := fillingConfirmButton);
cappingConfirmR(CLK := cappingConfirmButton);
packingConfirmR(CLK := packingConfirmButton);
finishedR(CLK := finishedButton);

Pump_Motor := FALSE;
Filling_Valve := FALSE;
Capping_Machine := FALSE;
Packing_Machine := FALSE;
Completion_Light := FALSE;

CASE State OF
    1:
        Pump_Motor := TRUE;
    2:
        Filling_Valve := TRUE;
    3:
        Capping_Machine := TRUE;
    4:
        Packing_Machine := TRUE;
    5:
        Completion_Light := TRUE;
END_CASE

IF State = 0 AND bottleSensorR.Q THEN
    State := 1;
ELSIF State = 1 AND cleaningConfirmR.Q THEN
    State := 2;
ELSIF State = 2 AND fillingConfirmR.Q THEN
    State := 3;
ELSIF State = 3 AND cappingConfirmR.Q THEN
    State := 4;
ELSIF State = 4 AND packingConfirmR.Q THEN
    State := 5;
ELSIF State = 5 AND finishedR.Q THEN
    State := 0;
END_IF

(* ---- public-easy-01.candidate_02.st ---- *)
PROGRAM FillingLineControl
VAR_INPUT
    bottleSensor : BOOL;
    cleaningConfirmButton : BOOL;
    fillingConfirmButton : BOOL;
    cappingConfirmButton : BOOL;
    packingConfirmButton : BOOL;
    finishedButton : BOOL;
END_VAR
VAR_OUTPUT
    Pump_Motor : BOOL;
    Filling_Valve : BOOL;
    Capping_Machine : BOOL;
    Packing_Machine : BOOL;
    Completion_Light : BOOL;
END_VAR
VAR
    State : INT := 0;
    bottleSensorR : R_TRIG;
    cleaningConfirmR : R_TRIG;
    fillingConfirmR : R_TRIG;
    cappingConfirmR : R_TRIG;
    packingConfirmR : R_TRIG;
    finishedR : R_TRIG;
END_VAR

bottleSensorR(CLK := bottleSensor);
cleaningConfirmR(CLK := cleaningConfirmButton);
fillingConfirmR(CLK := fillingConfirmButton);
cappingConfirmR(CLK := cappingConfirmButton);
packingConfirmR(CLK := packingConfirmButton);
finishedR(CLK := finishedButton);

Pump_Motor := FALSE;
Filling_Valve := FALSE;
Capping_Machine := FALSE;
Packing_Machine := FALSE;
Completion_Light := FALSE;

CASE State OF
    1:
        Pump_Motor := TRUE;
    2:
        Filling_Valve := TRUE;
    3:
        Capping_Machine := TRUE;
    4:
        Packing_Machine := TRUE;
    5:
        Completion_Light := TRUE;
END_CASE

IF State = 0 AND bottleSensorR.Q THEN
    State := 1;
ELSIF State = 1 AND cleaningConfirmR.Q THEN
    State := 2;
ELSIF State = 2 AND fillingConfirmR.Q THEN
    State := 3;
ELSIF State = 3 AND cappingConfirmR.Q THEN
    State := 4;
ELSIF State = 4 AND packingConfirmR.Q THEN
    State := 5;
ELSIF State = 5 AND finishedR.Q THEN
    State := 0;
END_IF

END_PROGRAM
